Fanuc KAREL source: kb00159.KL

-- PROVISIONAL review KL for V1013-1; original PC SHA256 5d484ac70e92e9c7b9312b77c14d3a1681a0e297d40bfb83b739b98c6ba181bb
-- Incomplete behavior may be omitted. Consult companion uncertainty JSON. Do not deploy.
PROGRAM KB00159
%NOLOCKGROUP
BEGIN
  -- UNRESOLVED_PC offsets 5-14; opcodes 3F,75
  -- UNRESOLVED_PC offsets 19-26; opcodes 9D,23
  -- UNRESOLVED_PC offsets 31-38; opcodes 9D,23
  -- UNRESOLVED_PC offsets 43-52; opcodes 3F,75
  -- UNRESOLVED_PC offsets 57-64; opcodes 9D,23
  -- UNRESOLVED_PC offsets 69-107; opcodes 27,22,2A,22,22,22,2A,22,31
  -- UNRESOLVED_PC offsets 112-116; opcodes 7F
END KB00159
